Fanuc KAREL source: KC00057.KL

PROGRAM KC00057
%NOLOCKGROUP
%ENVIRONMENT DEBUG
VAR
  I: INTEGER
  J: INTEGER
  K: INTEGER
  R: REAL
  B: BOOLEAN
  S: STRING[80]
  T: STRING[80]
  P: PATH
  Q: PATH
  AI: ARRAY[8] OF INTEGER
  AB: ARRAY[244] OF BYTE
BEGIN
  SET_DB_EVENT(I,B)
END KC00057
